// TIA Portal V21 export
VAR_GLOBAL   // PLC tag table "Conveyor I/O"
   Ib_CarrierPresent AT %I1300.3 : Bool;   // Carrier vorhanden / Carrier present   {ExternalAccessible false}
   Qr_Speed AT %QD40 : Real;
END_VAR
VAR_GLOBAL CONSTANT   // user constants
   MaxCarriers : Int := 12;   // Maximum carriers on the line
END_VAR
